Staubli VAL3: utLabel.dtx

public utAppearance Appearance
  [0]
    string sBackgroundColour
    string sColour
    bool bVisibility
public utBorder Border
  [0]
    string sBorderColour
    string sBorderStyle
    num nBorderWidth
public utCommon Common
  [0]
    string sText
    string sID
    string sPage
public utText Text
  [0]
    string sFontFamily
    string sFontStyle
    string sFontWeight
    string sTextAlignment
    num nFontSize
public utEvents Events
  [0]
    bool bClick
    bool bMouseDown
    bool bMouseUp
public utData Data
  [0]
    num nVal
    bool bStatus
